// TIA Portal V20 export
// export: Created 2026-10-12T15:52:20.8909765Z, ExportSetting WithDefaults, DisplayName Totally Integrated Automation Portal, DisplayVersion V20, DisplayName TIA Portal Openness, DisplayVersion V20, DisplayName TIA Portal Teamcenter Gateway, DisplayVersion V20, DisplayName TIA Portal Version Control Interface, DisplayVersion V20, DisplayName SINAMICS Startdrive Advanced, DisplayVersion V20 SP1 Update 2, DisplayName SINAMICS Startdrive G110M, G120, G120C, G120D, G120P, G115D, DisplayVersion V20 SP1 Update 2, DisplayName SINAMICS Startdrive G130, G150, S120, S150, SINAMICS MV, G220, S200, S210, DisplayVersion V20 SP1 Update 2, DisplayName STEP 7 Professional, DisplayVersion V20, DisplayName STEP 7 Safety, DisplayVersion V20, DisplayName WinCC Basic/Comfort/Advanced, DisplayVersion V20, DisplayName WinCC Professional, DisplayVersion V20, DisplayName WinCC Unified, DisplayVersion V20
FUNCTION "F_AlarmPersistenceBench" : Void   // FC175, SCL
{ S7_Optimized_Access := 'TRUE' }
VERSION : 0.1
// stored: AutoNumber true, IsIECCheckEnabled false, SetENOAutomatically false, UDAEnableTagReadback false
   VAR_TEMP
      Slot : Int;
      Index : Int;
      Text : WString[255];
      Symbol : WString[1];
   END_VAR
BEGIN

   #Slot := "FRK_AlarmHistoryIndex"(Scope := "GDB_AlarmPersistTest".Scope);
   "GDB_AlarmPersistTest".Slot := #Slot;
   IF #Slot < 1 THEN
       RETURN;
   END_IF;
   "GDB_AlarmPersistTest".Generation := "FRK_AlarmHistory".Rows[#Slot].Generation;
   "GDB_AlarmPersistTest".Checksum := "FRK_AlarmHistory".Rows[#Slot].Checksum;
   "GDB_AlarmPersistTest".Used := "FRK_AlarmHistory".Rows[#Slot].RingUsed;
   "GDB_AlarmPersistTest".Applied := "GDB_AlarmPersistTest".Operation <> 0;
   #Text := "GDB_AlarmPersistTest".Text;
   IF "GDB_AlarmPersistTest".UnicodeMode = 1 THEN
       #Symbol := WSTRING#' ';
       #Symbol[1] := UINT_TO_WCHAR(955);
       #Text := CONCAT(IN1 := #Text, IN2 := #Symbol);
       #Text := CONCAT(IN1 := #Text, IN2 := WSTRING#' ');
       #Symbol[1] := UINT_TO_WCHAR(20013);
       #Text := CONCAT(IN1 := #Text, IN2 := #Symbol);
   ELSIF "GDB_AlarmPersistTest".UnicodeMode = 2 THEN
       #Text := WSTRING#'';
       FOR #Index := 1 TO 85 DO
           #Symbol := WSTRING#' ';
           #Symbol[1] := UINT_TO_WCHAR(955);
           #Text := CONCAT(IN1 := #Text, IN2 := #Symbol);
           #Symbol[1] := UINT_TO_WCHAR(20013);
           #Text := CONCAT(IN1 := #Text, IN2 := #Symbol);
           #Text := CONCAT(IN1 := #Text, IN2 := WSTRING#'x');
       END_FOR;
   END_IF;
   CASE "GDB_AlarmPersistTest".Operation OF
       1, 2:
           IF "GDB_AlarmPersistTest".Scope = 'StationA' THEN
               IF "GDB_AlarmPersistTest".Operation = 1 THEN
                   "FRK_AlarmMessage"(Reason := "GDB_AlarmPersistTest".Reason,
                                      Description := #Text,
                                      SourcePath := WSTRING#'StationA',
                                      AlarmLog := "StationA".AlarmLog);
               ELSE
                   "FRK_AlarmBegin"(Startup := TRUE,
                                    AlarmLog := "StationA".AlarmLog);
               END_IF;
           END_IF;
           IF "GDB_AlarmPersistTest".Scope = 'StationA.Satellite' THEN
               IF "GDB_AlarmPersistTest".Operation = 1 THEN
                   "FRK_AlarmMessage"(Reason := "GDB_AlarmPersistTest".Reason,
                                      Description := #Text,
                                      SourcePath := WSTRING#'StationA.Satellite',
                                      AlarmLog := "StationA".Satellite.AlarmLog);
               ELSE
                   "FRK_AlarmBegin"(Startup := TRUE,
                                    AlarmLog := "StationA".Satellite.AlarmLog);
               END_IF;
           END_IF;
           IF "GDB_AlarmPersistTest".Scope = 'StationA.Satellite.Inner' THEN
               IF "GDB_AlarmPersistTest".Operation = 1 THEN
                   "FRK_AlarmMessage"(Reason := "GDB_AlarmPersistTest".Reason,
                                      Description := #Text,
                                      SourcePath := WSTRING#'StationA.Satellite.Inner',
                                      AlarmLog := "StationA".Satellite.Inner.AlarmLog);
               ELSE
                   "FRK_AlarmBegin"(Startup := TRUE,
                                    AlarmLog := "StationA".Satellite.Inner.AlarmLog);
               END_IF;
           END_IF;
           IF "GDB_AlarmPersistTest".Scope = 'StationB' THEN
               IF "GDB_AlarmPersistTest".Operation = 1 THEN
                   "FRK_AlarmMessage"(Reason := "GDB_AlarmPersistTest".Reason,
                                      Description := #Text,
                                      SourcePath := WSTRING#'StationB',
                                      AlarmLog := "StationB".AlarmLog);
               ELSE
                   "FRK_AlarmBegin"(Startup := TRUE,
                                    AlarmLog := "StationB".AlarmLog);
               END_IF;
           END_IF;
           IF "GDB_AlarmPersistTest".Scope = 'StationB.Satellite' THEN
               IF "GDB_AlarmPersistTest".Operation = 1 THEN
                   "FRK_AlarmMessage"(Reason := "GDB_AlarmPersistTest".Reason,
                                      Description := #Text,
                                      SourcePath := WSTRING#'StationB.Satellite',
                                      AlarmLog := "StationB".Satellite.AlarmLog);
               ELSE
                   "FRK_AlarmBegin"(Startup := TRUE,
                                    AlarmLog := "StationB".Satellite.AlarmLog);
               END_IF;
           END_IF;
           IF "GDB_AlarmPersistTest".Scope = 'StationB.Satellite.Inner' THEN
               IF "GDB_AlarmPersistTest".Operation = 1 THEN
                   "FRK_AlarmMessage"(Reason := "GDB_AlarmPersistTest".Reason,
                                      Description := #Text,
                                      SourcePath := WSTRING#'StationB.Satellite.Inner',
                                      AlarmLog := "StationB".Satellite.Inner.AlarmLog);
               ELSE
                   "FRK_AlarmBegin"(Startup := TRUE,
                                    AlarmLog := "StationB".Satellite.Inner.AlarmLog);
               END_IF;
           END_IF;
       10:
           "FRK_AlarmHistory".Rows[#Slot].SchemaVersion := 2;
       11:
           "FRK_AlarmHistory".Rows[#Slot].RingHead := 65;
       12:
           "FRK_AlarmHistory".Rows[#Slot].Checksum := "FRK_AlarmHistory".Rows[#Slot].Checksum XOR DWORD#1;
       13:
           "FRK_AlarmHistory".Rows[#Slot].Scope := 'foreign';
       14:
           "FRK_AlarmHistory".Rows[#Slot].Ring[1].Description := WSTRING#'corrupted';
       15:
           "FRK_AlarmHistory".Rows[#Slot].Ring[1].Duration := T#-1ms;
       16:
           "FRK_AlarmHistory".Rows[#Slot].SchemaVersion := 0;
           "FRK_AlarmHistory".Rows[#Slot].Generation := 0;
           "FRK_AlarmHistory".Rows[#Slot].Scope := '';
           "FRK_AlarmHistory".Rows[#Slot].Checksum := DWORD#0;
       17:
           "FRK_AlarmHistory".Rows[#Slot].RingUsed := -1;
   END_CASE;
   "GDB_AlarmPersistTest".Operation := 0;
END_FUNCTION
